(* IEC 61131-3 sources: Repository_IEMA_Test/LMC_PacDrive.device.xml.v3^/Plc Logic.plclogic.xml.v3^/Application.application.xml.v3^/TemplateFullProgrammingFramework/Examples/ExampleDiagSources/FB_ExampleTableDiagSource.fb.st^, 6 files *)

(* ---- CancelWriting.meth.st ---- *)
{attribute 'hide'}
METHOD CancelWriting : BOOL
VAR_INPUT
END_VAR

(* Deactivate writing if we are (for whatever reason) no longer adressed.
   May happen in case network connection with Diagnostics is disrupted or Source will be disabled *)

THIS^.diOldCmd			:= 0;
THIS^.diCmdExecState	:= 0;

(* ---- DiagQuit.meth.st ---- *)
{attribute 'hide'}
METHOD DiagQuit : BOOL
VAR_INPUT
END_VAR

IF THIS^.i_xEnable AND THIS^.q_xActive AND THIS^.q_etDiag <> GD.ET_Diag.Ok AND THIS^.diState = 0 THEN

	THIS^.rtrigDiagQuit(CLK := THIS^.i_xDiagQuit);
	IF THIS^.rtrigDiagQuit.Q THEN
		CancelWriting();

		THIS^.udiOwnSourceId	:= 0;

		THIS^.fbTableWriter.FB_Init(bInitRetains := FALSE, bInCopyCode := FALSE);

		THIS^.q_xReady		:= TRUE;
		THIS^.q_etDiag		:= GD.ET_Diag.Ok;
		THIS^.q_etDiagExt	:= ET_DiagExt.WaitUntilDiagnosticsManagerReady;
		THIS^.q_sMsg		:= '';

		THIS^.diState := 10;
	END_IF

END_IF

(* ---- ExceptionDuringWriting.meth.st ---- *)
{attribute 'hide'}
METHOD ExceptionDuringWriting : BOOL
VAR_INPUT
END_VAR

(* exception during writing *)
CASE THIS^.etDiagExtTPL OF
	TPL.ET_DiagExt.HeaderStartAlreadySuccessfullyCalled,	// FB_TableWriter.HeaderStart
	TPL.ET_DiagExt.FileIdNotSet,							// FB_TableWriter.HeaderStart
	TPL.ET_DiagExt.FileIdInvalid,							// FB_TableWriter.HeaderStart & FB_TableWriter.HeaderAddColumn & FB_TableWriter.HeaderFinish & FB_TableWriter.RowStart & FB_TableWriter.RowValue & FB_TableWriter.TableEnd
	TPL.ET_DiagExt.FileNotOpen,								// FB_TableWriter.HeaderStart & FB_TableWriter.HeaderAddColumn & FB_TableWriter.HeaderFinish & FB_TableWriter.RowStart & FB_TableWriter.RowValue & FB_TableWriter.TableEnd
	TPL.ET_DiagExt.UnexpectedFeedback,						// FB_TableWriter.HeaderStart & FB_TableWriter.HeaderAddColumn & FB_TableWriter.HeaderFinish & FB_TableWriter.RowStart & FB_TableWriter.RowValue & FB_TableWriter.TableEnd
	TPL.ET_DiagExt.HeaderStartNotCalled,					// FB_TableWriter.HeaderAddColumn
	TPL.ET_DiagExt.HeaderStartNotSuccessfullyCalled,		// FB_TableWriter.HeaderAddColumn
	TPL.ET_DiagExt.MaxNumberOfColumnsExceeded,				// FB_TableWriter.HeaderAddColumn
	TPL.ET_DiagExt.NameInvalid,								// FB_TableWriter.HeaderAddColumn
	TPL.ET_DiagExt.NoColumnsDefined,						// FB_TableWriter.HeaderFinish
	TPL.ET_DiagExt.DefineHeaderFirst,						// FB_TableWriter.RowStart
	TPL.ET_DiagExt.RowStartedCallRowEndFirst,				// FB_TableWriter.RowStart
	TPL.ET_DiagExt.CallRowStartFirst,						// FB_TableWriter.RowValue
	TPL.ET_DiagExt.ColumnNumberRange,						// FB_TableWriter.RowValue
	TPL.ET_DiagExt.RowsStillOpen,							// FB_TableWriter.TableEnd
	TPL.ET_DiagExt.HeaderColumnIdInvalid:

		SetDiagOutputs(	i_etDiag	:= GD.ET_Diag.UnexpectedProgramBehavior,
						i_etDiagExt	:= ET_DiagExt.UnexpectedFeedback,
						i_sMsg		:= PDL.FC_MultiConcat(	i_sString1	:= 'FB_TableWriter: ',
															i_sString2	:= GD.FC_EtDiagToString(THIS^.etDiag),
															i_sString3	:= ' - ',
															i_sString4	:= TPL.FC_EtDiagExtToString(THIS^.etDiagExtTPL),
															q_etDiag	=> ,
															q_etDiagExt	=> ));
	ELSE
		SetDiagOutputs(	i_etDiag	:= GD.ET_Diag.UnexpectedProgramBehavior,
						i_etDiagExt	:= ET_DiagExt.UnexpectedFeedback,
						i_sMsg		:= PDL.FC_MultiConcat(	i_sString1	:= 'FB_TableWriter: ',
															i_sString2	:= GD.FC_EtDiagToString(THIS^.etDiag),
															i_sString3	:= ' - ',
															i_sString4	:= TPL.FC_EtDiagExtToString(THIS^.etDiagExtTPL),
															q_etDiag	=> ,
															q_etDiagExt	=> ));
END_CASE

CancelWriting();

(* ---- SetDiagOutputs.meth.st ---- *)
{attribute 'hide'}
METHOD SetDiagOutputs : BOOL
VAR_INPUT
	i_etDiag		: GD.ET_Diag;
	i_etDiagExt		: ET_DiagExt;
	i_sMsg			: STRING[80];
END_VAR

IF THIS^.q_etDiag = GD.ET_Diag.Ok OR i_etDiagExt = ET_DiagExt.Disabled THEN

	IF i_etDiag <> GD.ET_Diag.Ok OR i_etDiagExt = ET_DiagExt.Disabled THEN

		IF i_etDiag <> GD.ET_Diag.Ok THEN
			THIS^.iq_stComStructure.iq_diCmd := -THIS^.iq_stComStructure.iq_diCmd;
		END_IF

		IF i_etDiagExt = ET_DiagExt.Disabled THEN
			THIS^.q_xActive := FALSE;

			CancelWriting();
		END_IF

		THIS^.q_xReady := FALSE;
		THIS^.diState := 0;
	END_IF

	THIS^.q_etDiag		:= i_etDiag;
	THIS^.q_etDiagExt	:= i_etDiagExt;
	THIS^.q_sMsg		:= i_sMsg;

END_IF

(* ---- WriteDiagDataControl.meth.st ---- *)
{attribute 'hide'}
METHOD WriteDiagDataControl : BOOL
VAR_INPUT
END_VAR

IF (THIS^.diOldCmd <> THIS^.iq_stComStructure.iq_diCmd AND THIS^.iq_stComStructure.iq_diCmd > 0) THEN

	THIS^.diOldCmd := THIS^.iq_stComStructure.iq_diCmd;

	(* new command, start execution *)
	CASE THIS^.iq_stComStructure.iq_diCmd OF

		1: (* write diag data to file *)
			IF (THIS^.iq_stComStructure.i_diFileId > 0) THEN

				SetDiagOutputs(	i_etDiag		:= GD.ET_Diag.Ok,
								i_etDiagExt		:= ET_DiagExt.WritingToFile,
								i_sMsg			:= '');

				THIS^.iq_stComStructure.q_lrProgress := 0.0;

				THIS^.fbTableWriter.diFileId := THIS^.iq_stComStructure.i_diFileId;

				THIS^.diCmdExecState := 1; (* start writing to file *)
			ELSE
				(* invalid file id *)
				SetDiagOutputs(	i_etDiag		:= GD.ET_Diag.InputParameterInvalid,
								i_etDiagExt		:= ET_DiagExt.FileIdInvalid,
								i_sMsg			:= CONCAT('Invalid file Id iq_stComStructure.i_diFileId: ', DINT_TO_STRING(THIS^.iq_stComStructure.i_diFileId)));
			END_IF
		ELSE
			(* unkown cmd *)
			SetDiagOutputs(	i_etDiag		:= GD.ET_Diag.InputParameterInvalid,
							i_etDiagExt		:= ET_DiagExt.CmdUnknown,
							i_sMsg			:= CONCAT('Unknown command iq_stComStructure.diCmd: ', DINT_TO_STRING(THIS^.iq_stComStructure.iq_diCmd)));

			CancelWriting();
	END_CASE
END_IF

(* ---- WriteDiagDataToFile.meth.st ---- *)
{attribute 'hide'}
METHOD WriteDiagDataToFile : BOOL
VAR_INPUT
END_VAR

TPL.FC_CanContinueWriting(iq_stCanContinueWriting := THIS^.iq_stComStructure.iq_stCanContinueWriting); (* loop as long as we can continue to write *)

WHILE (THIS^.iq_stComStructure.iq_stCanContinueWriting.xCanContinue) DO

	CASE THIS^.diCmdExecState OF
		1:
			(* start writing *)
			THIS^.fbTableWriter.HeaderStart(	i_sName					:= THIS^.c_sName,
												i_sTypeName				:= THIS^.c_sTypeName,
												i_sTitleEnglish			:= 'Example Data as Table',
												i_sTitleGerman			:= 'Beispieldaten als Tabelle',
												i_uiPrintRank			:= 14,
												i_sEmptyListTextEnglish	:= 'No data available to show',
												i_sEmptyListTextGerman	:= 'Keine Daten zum Anzeigen vorhanden',
												q_etDiag				=> THIS^.etDiag,
												q_etDiagExt				=> THIS^.etDiagExtTPL);

			IF THIS^.etDiag <> GD.ET_Diag.Ok THEN
				ExceptionDuringWriting();
				EXIT;
			END_IF

			THIS^.udiCName := THIS^.fbTableWriter.HeaderAddColumn(	i_sName			:= 'Name',
																	i_sTextEnglish	:= 'Name',
																	i_sTextGerman	:= 'Name',
																	i_uiWidth		:= 120,
																	q_etDiag		=> THIS^.etDiag,
																	q_etDiagExt		=> THIS^.etDiagExtTPL);
			IF THIS^.etDiag <> GD.ET_Diag.Ok THEN
				ExceptionDuringWriting();
				EXIT;
			END_IF

			THIS^.udiCValue := THIS^.fbTableWriter.HeaderAddColumn(	i_sName			:= 'Value',
																	i_sTextEnglish	:= 'Value',
																	i_sTextGerman	:= 'Wert',
																	i_uiWidth		:= 120,
																	q_etDiag		=> THIS^.etDiag,
																	q_etDiagExt		=> THIS^.etDiagExtTPL);
			IF THIS^.etDiag <> GD.ET_Diag.Ok THEN
				ExceptionDuringWriting();
				EXIT;
			END_IF

			THIS^.udiCC3 := THIS^.fbTableWriter.HeaderAddColumn(i_sName			:= 'Column3',
																i_sTextEnglish	:= 'Column3',
																i_sTextGerman	:= 'Spalte3',
																i_uiWidth		:= 120,
																q_etDiag		=> THIS^.etDiag,
																q_etDiagExt		=> THIS^.etDiagExtTPL);
			IF THIS^.etDiag <> GD.ET_Diag.Ok THEN
				ExceptionDuringWriting();
				EXIT;
			END_IF

			IF THIS^.udiCC3 <= 0 OR THIS^.udiCValue <= 0 OR THIS^.udiCName <= 0 THEN

				THIS^.etDiag		:= GD.ET_Diag.ExecutionAborted;
				THIS^.etDiagExtTPL	:= TPL.ET_DiagExt.HeaderColumnIdInvalid;

				ExceptionDuringWriting();
				EXIT;
			END_IF

			THIS^.fbTableWriter.HeaderFinish(	q_etDiag	=> THIS^.etDiag,
												q_etDiagExt	=> THIS^.etDiagExtTPL);

			IF THIS^.etDiag <> GD.ET_Diag.Ok THEN
				ExceptionDuringWriting();
				EXIT;
			END_IF

			THIS^.udiRowCounter := 1; (* start loop at index 1 *)

			THIS^.diCmdExecState := THIS^.diCmdExecState + 1;

		2:	(* loop over all rows *)

			IF (THIS^.udiRowCounter <= THIS^.c_udiMaxNumRows) THEN

				(* write row *)
				THIS^.fbTableWriter.RowStart(	q_etDiag	=> THIS^.etDiag,
												q_etDiagExt	=> THIS^.etDiagExtTPL);

				IF THIS^.etDiag <> GD.ET_Diag.Ok THEN
					ExceptionDuringWriting();
					EXIT;
				END_IF

				(* write values *)
				THIS^.fbTableWriter.RowValue(	i_udiColumnNumber	:= THIS^.udiCName,
												i_sValue			:= CONCAT('name_',UDINT_TO_STRING(udiRowCounter)),
												q_etDiag			=> THIS^.etDiag,
												q_etDiagExt			=> THIS^.etDiagExtTPL);

				IF THIS^.etDiag <> GD.ET_Diag.Ok THEN
					ExceptionDuringWriting();
					EXIT;
				END_IF

				THIS^.fbTableWriter.RowValue(	i_udiColumnNumber	:= THIS^.udiCValue,
												i_sValue			:= LREAL_TO_STRING((8000.0 - UDINT_TO_LREAL(udiRowCounter))/5),
												q_etDiag			=> THIS^.etDiag,
												q_etDiagExt			=> THIS^.etDiagExtTPL);

				IF THIS^.etDiag <> GD.ET_Diag.Ok THEN
					ExceptionDuringWriting();
					EXIT;
				END_IF

				THIS^.fbTableWriter.RowValue(	i_udiColumnNumber	:= THIS^.udiCC3,
												i_sValue			:= UDINT_TO_STRING(udiRowCounter + 88),
												q_etDiag			=> THIS^.etDiag,
												q_etDiagExt			=> THIS^.etDiagExtTPL);

				IF THIS^.etDiag <> GD.ET_Diag.Ok THEN
					ExceptionDuringWriting();
					EXIT;
				END_IF

				THIS^.fbTableWriter.RowEnd(	q_etDiag	=> THIS^.etDiag,
											q_etDiagExt	=> THIS^.etDiagExtTPL);

				IF THIS^.etDiag <> GD.ET_Diag.Ok THEN
					ExceptionDuringWriting();
					EXIT;
				END_IF
			END_IF

			THIS^.iq_stComStructure.q_lrProgress := UDINT_TO_LREAL(THIS^.udiRowCounter) * LREAL#100.0 / MAX(UDINT_TO_LREAL(THIS^.c_udiMaxNumRows), LREAL#0.0001);

			THIS^.udiRowCounter := THIS^.udiRowCounter + 1;
			IF (THIS^.udiRowCounter > THIS^.c_udiMaxNumRows) THEN
				(* loop over all rows done *)
				THIS^.diCmdExecState := THIS^.diCmdExecState + 1;
			END_IF
		3:
			THIS^.fbTableWriter.TableEnd(	q_etDiag	=> THIS^.etDiag,
											q_etDiagExt	=> THIS^.etDiagExtTPL);

			IF THIS^.etDiag <> GD.ET_Diag.Ok THEN
				ExceptionDuringWriting();
				EXIT;
			END_IF

			(* done *)
			THIS^.iq_stComStructure.iq_diCmd := 0;

			SetDiagOutputs(	i_etDiag	:= GD.ET_Diag.Ok,
							i_etDiagExt	:= ET_DiagExt.DataSuccessfullyWritten,
							i_sMsg		:= '');

			THIS^.diCmdExecState := 0;
			EXIT; (* exit the while loop *)
	END_CASE

	(* check again whether we can continue writing *)
	TPL.FC_CanContinueWriting(iq_stCanContinueWriting := THIS^.iq_stComStructure.iq_stCanContinueWriting);
END_WHILE
